Staubli VAL3: click_Start.pgx

program click_Start()
  local bool l_bResult
begin
  //启动机器人
  l_bResult=userPageConfirm("确认启动机器人？")
  if l_bResult
    rs:bToStartCycle=true
    delay(0.2)
    rs:bToStartCycle=false
  endIf
end
